(* IEC 61131-3 sources: kns-port-domestic/tools/plcopen/tests/fixtures/constructs/src/POUs/F_Clamp, 2 files *)

(* ---- F_Clamp.decl.st ---- *)
// Назначение: ограничение значения диапазоном [rMin, rMax]; при rMin > rMax границы меняются местами
// Автор:      <ИМЯ ФАМИЛИЯ>
// Версия:     0.1.0
// Документ:   docs/plcopen.md
FUNCTION F_Clamp : REAL
VAR_INPUT
    rValue : REAL;      // значение
    rMin : REAL;        // нижняя граница
    rMax : REAL;        // верхняя граница
END_VAR
VAR
    rLow : REAL;
    rHigh : REAL;
END_VAR

(* ---- F_Clamp.impl.st ---- *)
// границы в правильном порядке
IF rMin <= rMax THEN
    rLow := rMin;
    rHigh := rMax;
ELSE
    rLow := rMax;
    rHigh := rMin;
END_IF
F_Clamp := LIMIT(rLow, rValue, rHigh);
